// TIA Portal V20 export
// export: Created 2026-10-19T18:01:59.2377084Z, ExportSetting WithDefaults, DisplayName Totally Integrated Automation Portal, DisplayVersion V20 Update 6, DisplayName TIA Portal Openness, DisplayVersion V20 Update 6, DisplayName TIA Portal Version Control Interface, DisplayVersion V20 Update 6, DisplayName SINAMICS Startdrive Advanced, DisplayVersion V20 SP1, DisplayName SINAMICS Startdrive G130, G150, S120, S150, SINAMICS MV, G220, S200, S210, DisplayVersion V20 SP1, DisplayName SINAMICS Startdrive G110M, G120, G120C, G120D, G120P, G115D, DisplayVersion V20 SP1, DisplayName STEP 7 Professional, DisplayVersion V20 Update 6, DisplayName STEP 7 Safety, DisplayVersion V20 Update 2, DisplayName WinCC Basic/Comfort/Advanced, DisplayVersion V20 Update 6, DisplayName WinCC Unified, DisplayVersion V20 Update 6
ORGANIZATION_BLOCK "Main"   // OB1, LAD, ProgramCycle
TITLE = "Main Program Sweep (Cycle)"
{ S7_Optimized_Access := 'TRUE' }
VERSION : 0.1
// stored: AutoNumber true, IsIECCheckEnabled false, SetENOAutomatically false
   VAR_INPUT
      Initial_Call : Bool;   // Initial call of this OB
      Remanence : Bool;   // =True, if remanent data are available
   END_VAR
   VAR_TEMP   // added for the SCL form of the ladder/FBD networks
      _w1 : Bool;
      _w2 : Bool;
      _w3 : Bool;
      _w4 : Bool;
      _w5 : Bool;
   END_VAR
BEGIN

REGION Network 1: Communication
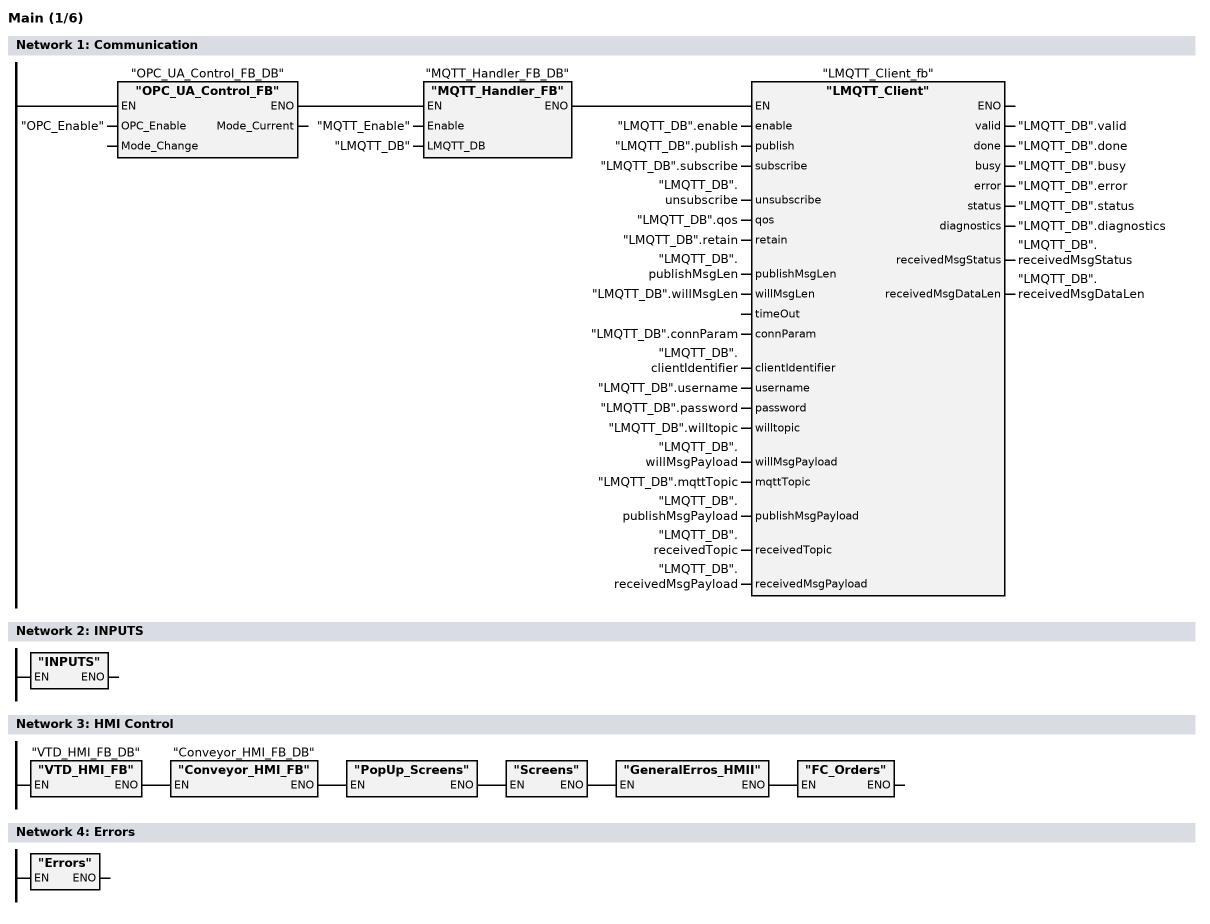
   RUNG wire#powerrail
      "OPC_UA_Control_FB_DB"(OPC_Enable := "OPC_Enable", Mode_Change :=, Mode_Current =>)
      "MQTT_Handler_FB_DB"(Enable := "MQTT_Enable", LMQTT_DB := "LMQTT_DB")
      "LMQTT_Client_fb"(enable := "LMQTT_DB".enable, publish := "LMQTT_DB".publish, subscribe := "LMQTT_DB".subscribe, unsubscribe := "LMQTT_DB".unsubscribe, qos := "LMQTT_DB".qos, retain := "LMQTT_DB".retain, publishMsgLen := "LMQTT_DB".publishMsgLen, willMsgLen := "LMQTT_DB".willMsgLen, timeOut :=, connParam := "LMQTT_DB".connParam, clientIdentifier := "LMQTT_DB".clientIdentifier, username := "LMQTT_DB".username, password := "LMQTT_DB".password, willtopic := "LMQTT_DB".willtopic, willMsgPayload := "LMQTT_DB".willMsgPayload, mqttTopic := "LMQTT_DB".mqttTopic, publishMsgPayload := "LMQTT_DB".publishMsgPayload, receivedTopic := "LMQTT_DB".receivedTopic, receivedMsgPayload := "LMQTT_DB".receivedMsgPayload, valid => "LMQTT_DB".valid, done => "LMQTT_DB".done, busy => "LMQTT_DB".busy, error => "LMQTT_DB".error, status => "LMQTT_DB".status, diagnostics => "LMQTT_DB".diagnostics, receivedMsgStatus => "LMQTT_DB".receivedMsgStatus, receivedMsgDataLen => "LMQTT_DB".receivedMsgDataLen)
   END_RUNG
   // the same network as SCL:
   "OPC_UA_Control_FB_DB"(OPC_Enable := "OPC_Enable", ENO => #_w1);   // "OPC_UA_Control_FB"
   "MQTT_Handler_FB_DB"(EN := #_w1, Enable := "MQTT_Enable", LMQTT_DB := "LMQTT_DB", ENO => #_w2);   // "MQTT_Handler_FB"
   IF #_w2 THEN
       "LMQTT_Client_fb"(enable := "LMQTT_DB".enable,   // "LMQTT_Client"
                         publish := "LMQTT_DB".publish,
                         subscribe := "LMQTT_DB".subscribe,
                         unsubscribe := "LMQTT_DB".unsubscribe,
                         qos := "LMQTT_DB".qos,
                         retain := "LMQTT_DB".retain,
                         publishMsgLen := "LMQTT_DB".publishMsgLen,
                         willMsgLen := "LMQTT_DB".willMsgLen,
                         connParam := "LMQTT_DB".connParam,
                         clientIdentifier := "LMQTT_DB".clientIdentifier,
                         username := "LMQTT_DB".username,
                         password := "LMQTT_DB".password,
                         willtopic := "LMQTT_DB".willtopic,
                         willMsgPayload := "LMQTT_DB".willMsgPayload,
                         mqttTopic := "LMQTT_DB".mqttTopic,
                         publishMsgPayload := "LMQTT_DB".publishMsgPayload,
                         receivedTopic := "LMQTT_DB".receivedTopic,
                         receivedMsgPayload := "LMQTT_DB".receivedMsgPayload,
                         valid => "LMQTT_DB".valid,
                         done => "LMQTT_DB".done,
                         busy => "LMQTT_DB".busy,
                         error => "LMQTT_DB".error,
                         status => "LMQTT_DB".status,
                         diagnostics => "LMQTT_DB".diagnostics,
                         receivedMsgStatus => "LMQTT_DB".receivedMsgStatus,
                         receivedMsgDataLen => "LMQTT_DB".receivedMsgDataLen);
   END_IF;
END_REGION

REGION Network 2: INPUTS
   RUNG wire#powerrail
      "INPUTS"()
   END_RUNG
   // the same network as SCL:
   "INPUTS"();
END_REGION

REGION Network 3: HMI Control
   RUNG wire#powerrail
      "VTD_HMI_FB_DB"()
      "Conveyor_HMI_FB_DB"()
      "PopUp_Screens"()
      "Screens"()
      "GeneralErros_HMII"()
      "FC_Orders"()
   END_RUNG
   // the same network as SCL:
   "VTD_HMI_FB_DB"(ENO => #_w1);   // "VTD_HMI_FB"
   "Conveyor_HMI_FB_DB"(EN := #_w1, ENO => #_w2);   // "Conveyor_HMI_FB"
   "PopUp_Screens"(EN := #_w2, ENO => #_w3);
   "Screens"(EN := #_w3, ENO => #_w4);
   "GeneralErros_HMII"(EN := #_w4, ENO => #_w5);
   IF #_w5 THEN "FC_Orders"(); END_IF;
END_REGION

REGION Network 4: Errors
   RUNG wire#powerrail
      "Errors"()
   END_RUNG
   // the same network as SCL:
   "Errors"();
END_REGION

REGION Network 5: Carousel Conveyors
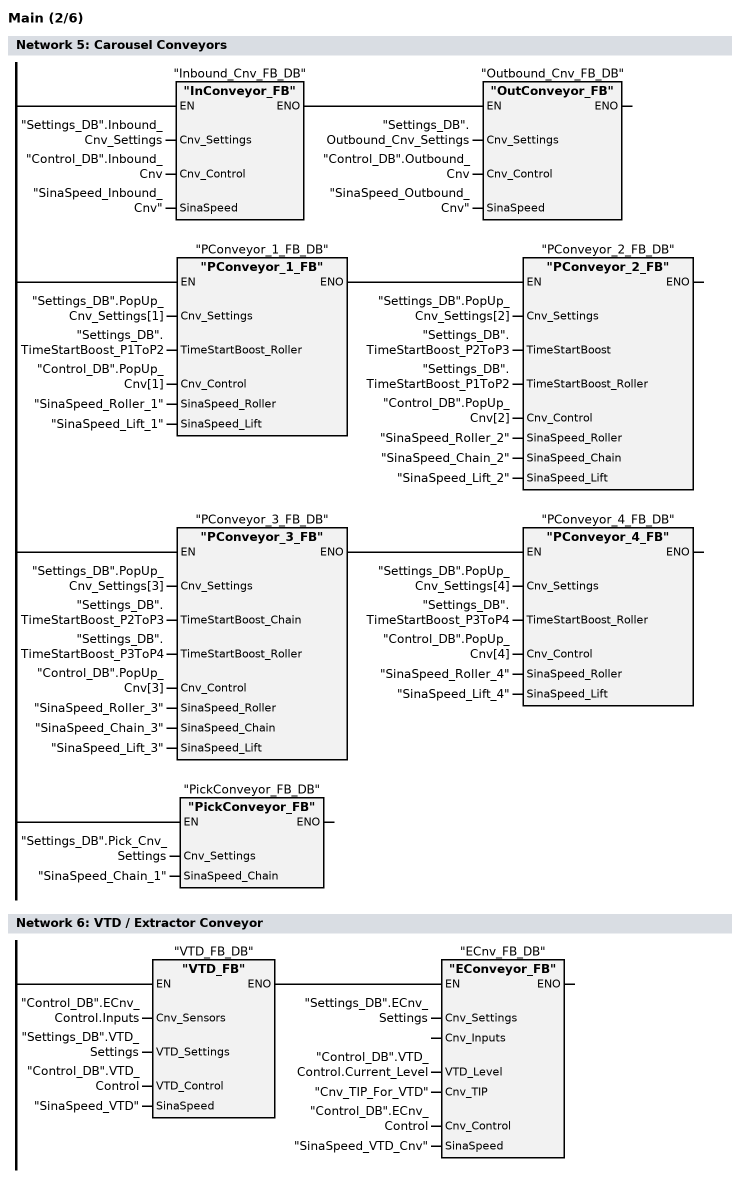
   RUNG wire#powerrail
      "Inbound_Cnv_FB_DB"(Cnv_Settings := "Settings_DB".Inbound_Cnv_Settings, Cnv_Control := "Control_DB".Inbound_Cnv, SinaSpeed := "SinaSpeed_Inbound_Cnv")
      "Outbound_Cnv_FB_DB"(Cnv_Settings := "Settings_DB".Outbound_Cnv_Settings, Cnv_Control := "Control_DB".Outbound_Cnv, SinaSpeed := "SinaSpeed_Outbound_Cnv")
   END_RUNG
   RUNG wire#powerrail
      "PConveyor_1_FB_DB"(Cnv_Settings := "Settings_DB".PopUp_Cnv_Settings[1], TimeStartBoost_Roller := "Settings_DB".TimeStartBoost_P1ToP2, Cnv_Control := "Control_DB".PopUp_Cnv[1], SinaSpeed_Roller := "SinaSpeed_Roller_1", SinaSpeed_Lift := "SinaSpeed_Lift_1")
      "PConveyor_2_FB_DB"(Cnv_Settings := "Settings_DB".PopUp_Cnv_Settings[2], TimeStartBoost := "Settings_DB".TimeStartBoost_P2ToP3, TimeStartBoost_Roller := "Settings_DB".TimeStartBoost_P1ToP2, Cnv_Control := "Control_DB".PopUp_Cnv[2], SinaSpeed_Roller := "SinaSpeed_Roller_2", SinaSpeed_Chain := "SinaSpeed_Chain_2", SinaSpeed_Lift := "SinaSpeed_Lift_2")
   END_RUNG
   RUNG wire#powerrail
      "PConveyor_3_FB_DB"(Cnv_Settings := "Settings_DB".PopUp_Cnv_Settings[3], TimeStartBoost_Chain := "Settings_DB".TimeStartBoost_P2ToP3, TimeStartBoost_Roller := "Settings_DB".TimeStartBoost_P3ToP4, Cnv_Control := "Control_DB".PopUp_Cnv[3], SinaSpeed_Roller := "SinaSpeed_Roller_3", SinaSpeed_Chain := "SinaSpeed_Chain_3", SinaSpeed_Lift := "SinaSpeed_Lift_3")
      "PConveyor_4_FB_DB"(Cnv_Settings := "Settings_DB".PopUp_Cnv_Settings[4], TimeStartBoost_Roller := "Settings_DB".TimeStartBoost_P3ToP4, Cnv_Control := "Control_DB".PopUp_Cnv[4], SinaSpeed_Roller := "SinaSpeed_Roller_4", SinaSpeed_Lift := "SinaSpeed_Lift_4")
   END_RUNG
   RUNG wire#powerrail
      "PickConveyor_FB_DB"(Cnv_Settings := "Settings_DB".Pick_Cnv_Settings, SinaSpeed_Chain := "SinaSpeed_Chain_1")
   END_RUNG
   // the same network as SCL:
   "Inbound_Cnv_FB_DB"(Cnv_Settings := "Settings_DB".Inbound_Cnv_Settings,   // "InConveyor_FB"
                       Cnv_Control := "Control_DB".Inbound_Cnv,
                       SinaSpeed := "SinaSpeed_Inbound_Cnv",
                       ENO => #_w1);
   IF #_w1 THEN
       "Outbound_Cnv_FB_DB"(Cnv_Settings := "Settings_DB".Outbound_Cnv_Settings,   // "OutConveyor_FB"
                            Cnv_Control := "Control_DB".Outbound_Cnv,
                            SinaSpeed := "SinaSpeed_Outbound_Cnv");
   END_IF;
   "PConveyor_1_FB_DB"(Cnv_Settings := "Settings_DB".PopUp_Cnv_Settings[1],   // "PConveyor_1_FB"
                       TimeStartBoost_Roller := "Settings_DB".TimeStartBoost_P1ToP2,
                       Cnv_Control := "Control_DB".PopUp_Cnv[1],
                       SinaSpeed_Roller := "SinaSpeed_Roller_1",
                       SinaSpeed_Lift := "SinaSpeed_Lift_1",
                       ENO => #_w2);
   IF #_w2 THEN
       "PConveyor_2_FB_DB"(Cnv_Settings := "Settings_DB".PopUp_Cnv_Settings[2],   // "PConveyor_2_FB"
                           TimeStartBoost := "Settings_DB".TimeStartBoost_P2ToP3,
                           TimeStartBoost_Roller := "Settings_DB".TimeStartBoost_P1ToP2,
                           Cnv_Control := "Control_DB".PopUp_Cnv[2],
                           SinaSpeed_Roller := "SinaSpeed_Roller_2",
                           SinaSpeed_Chain := "SinaSpeed_Chain_2",
                           SinaSpeed_Lift := "SinaSpeed_Lift_2");
   END_IF;
   "PConveyor_3_FB_DB"(Cnv_Settings := "Settings_DB".PopUp_Cnv_Settings[3],   // "PConveyor_3_FB"
                       TimeStartBoost_Chain := "Settings_DB".TimeStartBoost_P2ToP3,
                       TimeStartBoost_Roller := "Settings_DB".TimeStartBoost_P3ToP4,
                       Cnv_Control := "Control_DB".PopUp_Cnv[3],
                       SinaSpeed_Roller := "SinaSpeed_Roller_3",
                       SinaSpeed_Chain := "SinaSpeed_Chain_3",
                       SinaSpeed_Lift := "SinaSpeed_Lift_3",
                       ENO => #_w3);
   IF #_w3 THEN
       "PConveyor_4_FB_DB"(Cnv_Settings := "Settings_DB".PopUp_Cnv_Settings[4],   // "PConveyor_4_FB"
                           TimeStartBoost_Roller := "Settings_DB".TimeStartBoost_P3ToP4,
                           Cnv_Control := "Control_DB".PopUp_Cnv[4],
                           SinaSpeed_Roller := "SinaSpeed_Roller_4",
                           SinaSpeed_Lift := "SinaSpeed_Lift_4");
   END_IF;
   "PickConveyor_FB_DB"(Cnv_Settings := "Settings_DB".Pick_Cnv_Settings, SinaSpeed_Chain := "SinaSpeed_Chain_1");   // "PickConveyor_FB"
END_REGION

REGION Network 6: VTD / Extractor Conveyor
   RUNG wire#powerrail
      "VTD_FB_DB"(Cnv_Sensors := "Control_DB".ECnv_Control.Inputs, VTD_Settings := "Settings_DB".VTD_Settings, VTD_Control := "Control_DB".VTD_Control, SinaSpeed := "SinaSpeed_VTD")
      "ECnv_FB_DB"(Cnv_Settings := "Settings_DB".ECnv_Settings, Cnv_Inputs :=, VTD_Level := "Control_DB".VTD_Control.Current_Level, Cnv_TIP := "Cnv_TIP_For_VTD", Cnv_Control := "Control_DB".ECnv_Control, SinaSpeed := "SinaSpeed_VTD_Cnv")
   END_RUNG
   // the same network as SCL:
   "VTD_FB_DB"(Cnv_Sensors := "Control_DB".ECnv_Control.Inputs,   // "VTD_FB"
               VTD_Settings := "Settings_DB".VTD_Settings,
               VTD_Control := "Control_DB".VTD_Control,
               SinaSpeed := "SinaSpeed_VTD",
               ENO => #_w1);
   IF #_w1 THEN
       "ECnv_FB_DB"(Cnv_Settings := "Settings_DB".ECnv_Settings,   // "EConveyor_FB"
                    VTD_Level := "Control_DB".VTD_Control.Current_Level,
                    Cnv_TIP := "Cnv_TIP_For_VTD",
                    Cnv_Control := "Control_DB".ECnv_Control,
                    SinaSpeed := "SinaSpeed_VTD_Cnv");
   END_IF;
END_REGION

REGION Network 7: Level Conveyors
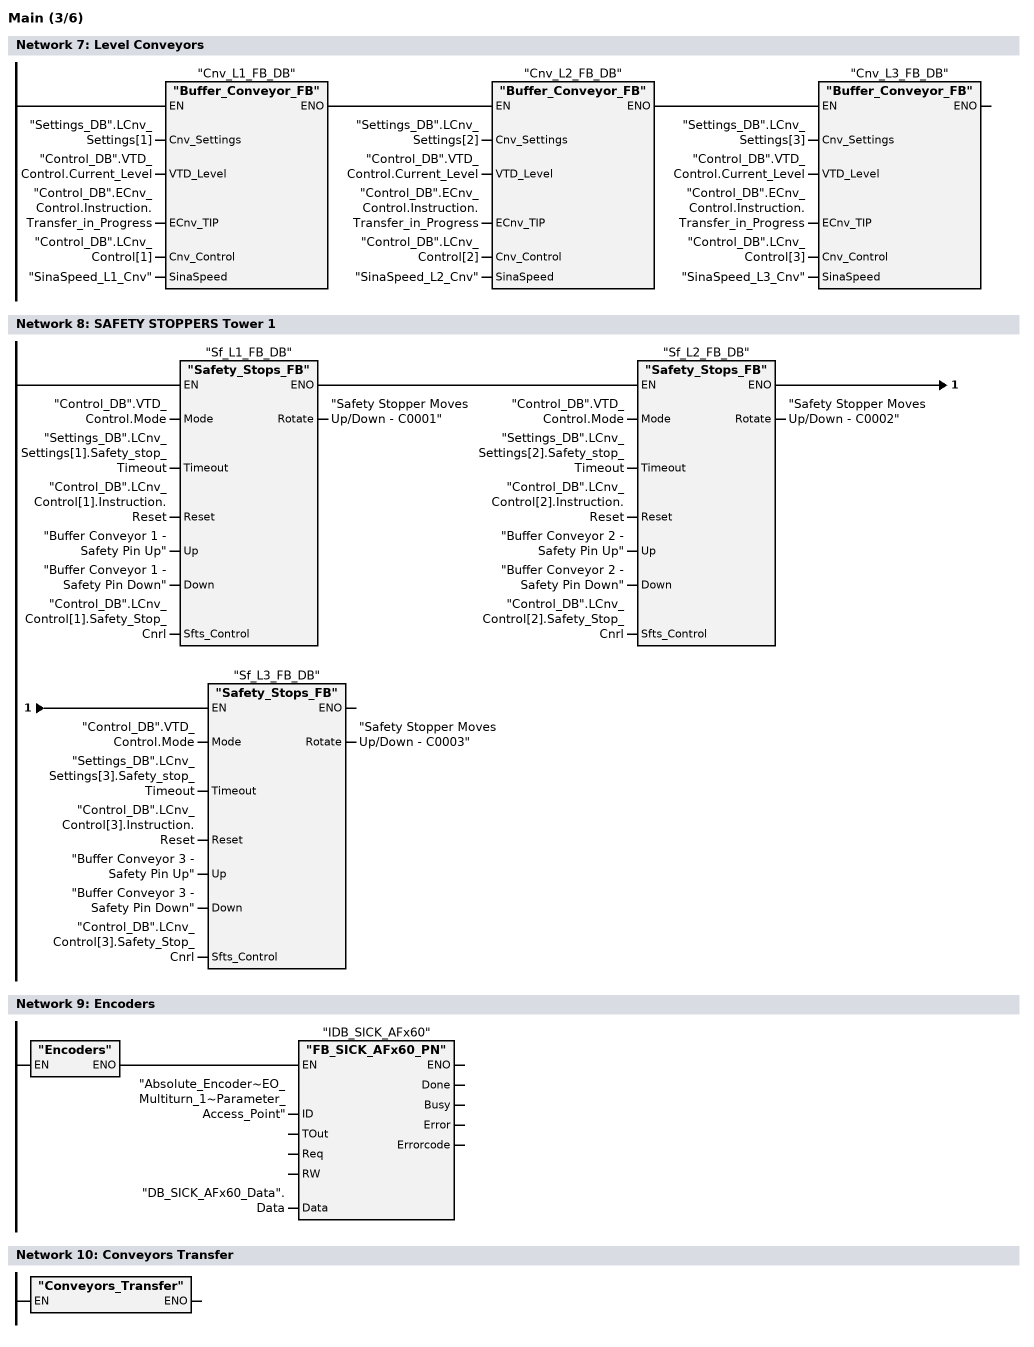
   RUNG wire#powerrail
      "Cnv_L1_FB_DB"(Cnv_Settings := "Settings_DB".LCnv_Settings[1], VTD_Level := "Control_DB".VTD_Control.Current_Level, ECnv_TIP := "Control_DB".ECnv_Control.Instruction.Transfer_in_Progress, Cnv_Control := "Control_DB".LCnv_Control[1], SinaSpeed := "SinaSpeed_L1_Cnv")
      "Cnv_L2_FB_DB"(Cnv_Settings := "Settings_DB".LCnv_Settings[2], VTD_Level := "Control_DB".VTD_Control.Current_Level, ECnv_TIP := "Control_DB".ECnv_Control.Instruction.Transfer_in_Progress, Cnv_Control := "Control_DB".LCnv_Control[2], SinaSpeed := "SinaSpeed_L2_Cnv")
      "Cnv_L3_FB_DB"(Cnv_Settings := "Settings_DB".LCnv_Settings[3], VTD_Level := "Control_DB".VTD_Control.Current_Level, ECnv_TIP := "Control_DB".ECnv_Control.Instruction.Transfer_in_Progress, Cnv_Control := "Control_DB".LCnv_Control[3], SinaSpeed := "SinaSpeed_L3_Cnv")
   END_RUNG
   // the same network as SCL:
   "Cnv_L1_FB_DB"(Cnv_Settings := "Settings_DB".LCnv_Settings[1],   // "Buffer_Conveyor_FB"
                  VTD_Level := "Control_DB".VTD_Control.Current_Level,
                  ECnv_TIP := "Control_DB".ECnv_Control.Instruction.Transfer_in_Progress,
                  Cnv_Control := "Control_DB".LCnv_Control[1],
                  SinaSpeed := "SinaSpeed_L1_Cnv",
                  ENO => #_w1);
   "Cnv_L2_FB_DB"(EN := #_w1,   // "Buffer_Conveyor_FB"
                  Cnv_Settings := "Settings_DB".LCnv_Settings[2],
                  VTD_Level := "Control_DB".VTD_Control.Current_Level,
                  ECnv_TIP := "Control_DB".ECnv_Control.Instruction.Transfer_in_Progress,
                  Cnv_Control := "Control_DB".LCnv_Control[2],
                  SinaSpeed := "SinaSpeed_L2_Cnv",
                  ENO => #_w2);
   IF #_w2 THEN
       "Cnv_L3_FB_DB"(Cnv_Settings := "Settings_DB".LCnv_Settings[3],   // "Buffer_Conveyor_FB"
                      VTD_Level := "Control_DB".VTD_Control.Current_Level,
                      ECnv_TIP := "Control_DB".ECnv_Control.Instruction.Transfer_in_Progress,
                      Cnv_Control := "Control_DB".LCnv_Control[3],
                      SinaSpeed := "SinaSpeed_L3_Cnv");
   END_IF;
END_REGION

REGION Network 8: SAFETY STOPPERS Tower 1
   RUNG wire#powerrail
      "Sf_L1_FB_DB"(Mode := "Control_DB".VTD_Control.Mode, Timeout := "Settings_DB".LCnv_Settings[1].Safety_stop_Timeout, Reset := "Control_DB".LCnv_Control[1].Instruction.Reset, Up := "Buffer Conveyor 1 - Safety Pin Up", Down := "Buffer Conveyor 1 - Safety Pin Down", Sfts_Control := "Control_DB".LCnv_Control[1].Safety_Stop_Cnrl, Rotate => "Safety Stopper Moves Up/Down - C0001")
      "Sf_L2_FB_DB"(Mode := "Control_DB".VTD_Control.Mode, Timeout := "Settings_DB".LCnv_Settings[2].Safety_stop_Timeout, Reset := "Control_DB".LCnv_Control[2].Instruction.Reset, Up := "Buffer Conveyor 2 - Safety Pin Up", Down := "Buffer Conveyor 2 - Safety Pin Down", Sfts_Control := "Control_DB".LCnv_Control[2].Safety_Stop_Cnrl, Rotate => "Safety Stopper Moves Up/Down - C0002")
      "Sf_L3_FB_DB"(Mode := "Control_DB".VTD_Control.Mode, Timeout := "Settings_DB".LCnv_Settings[3].Safety_stop_Timeout, Reset := "Control_DB".LCnv_Control[3].Instruction.Reset, Up := "Buffer Conveyor 3 - Safety Pin Up", Down := "Buffer Conveyor 3 - Safety Pin Down", Sfts_Control := "Control_DB".LCnv_Control[3].Safety_Stop_Cnrl, Rotate => "Safety Stopper Moves Up/Down - C0003")
   END_RUNG
   // the same network as SCL:
   "Sf_L1_FB_DB"(Mode := "Control_DB".VTD_Control.Mode,   // "Safety_Stops_FB"
                 Timeout := "Settings_DB".LCnv_Settings[1].Safety_stop_Timeout,
                 Reset := "Control_DB".LCnv_Control[1].Instruction.Reset,
                 Up := "Buffer Conveyor 1 - Safety Pin Up",
                 Down := "Buffer Conveyor 1 - Safety Pin Down",
                 Sfts_Control := "Control_DB".LCnv_Control[1].Safety_Stop_Cnrl,
                 Rotate => "Safety Stopper Moves Up/Down - C0001",
                 ENO => #_w1);
   "Sf_L2_FB_DB"(EN := #_w1,   // "Safety_Stops_FB"
                 Mode := "Control_DB".VTD_Control.Mode,
                 Timeout := "Settings_DB".LCnv_Settings[2].Safety_stop_Timeout,
                 Reset := "Control_DB".LCnv_Control[2].Instruction.Reset,
                 Up := "Buffer Conveyor 2 - Safety Pin Up",
                 Down := "Buffer Conveyor 2 - Safety Pin Down",
                 Sfts_Control := "Control_DB".LCnv_Control[2].Safety_Stop_Cnrl,
                 Rotate => "Safety Stopper Moves Up/Down - C0002",
                 ENO => #_w2);
   IF #_w2 THEN
       "Sf_L3_FB_DB"(Mode := "Control_DB".VTD_Control.Mode,   // "Safety_Stops_FB"
                     Timeout := "Settings_DB".LCnv_Settings[3].Safety_stop_Timeout,
                     Reset := "Control_DB".LCnv_Control[3].Instruction.Reset,
                     Up := "Buffer Conveyor 3 - Safety Pin Up",
                     Down := "Buffer Conveyor 3 - Safety Pin Down",
                     Sfts_Control := "Control_DB".LCnv_Control[3].Safety_Stop_Cnrl,
                     Rotate => "Safety Stopper Moves Up/Down - C0003");
   END_IF;
END_REGION

REGION Network 9: Encoders
   RUNG wire#powerrail
      "Encoders"()
      "IDB_SICK_AFx60"(ID := "Absolute_Encoder~EO_Multiturn_1~Parameter_Access_Point", TOut :=, Req :=, RW :=, Data := "DB_SICK_AFx60_Data".Data, Done =>, Busy =>, Error =>, Errorcode =>)
   END_RUNG
   // the same network as SCL:
   "Encoders"(ENO => #_w1);
   IF #_w1 THEN
       "IDB_SICK_AFx60"(ID := "Absolute_Encoder~EO_Multiturn_1~Parameter_Access_Point",   // "FB_SICK_AFx60_PN"
                        Data := "DB_SICK_AFx60_Data".Data);
   END_IF;
END_REGION

REGION Network 10: Conveyors Transfer
   RUNG wire#powerrail
      "Conveyors_Transfer"()
   END_RUNG
   // the same network as SCL:
   "Conveyors_Transfer"();
END_REGION

REGION Network 11: Lightbar
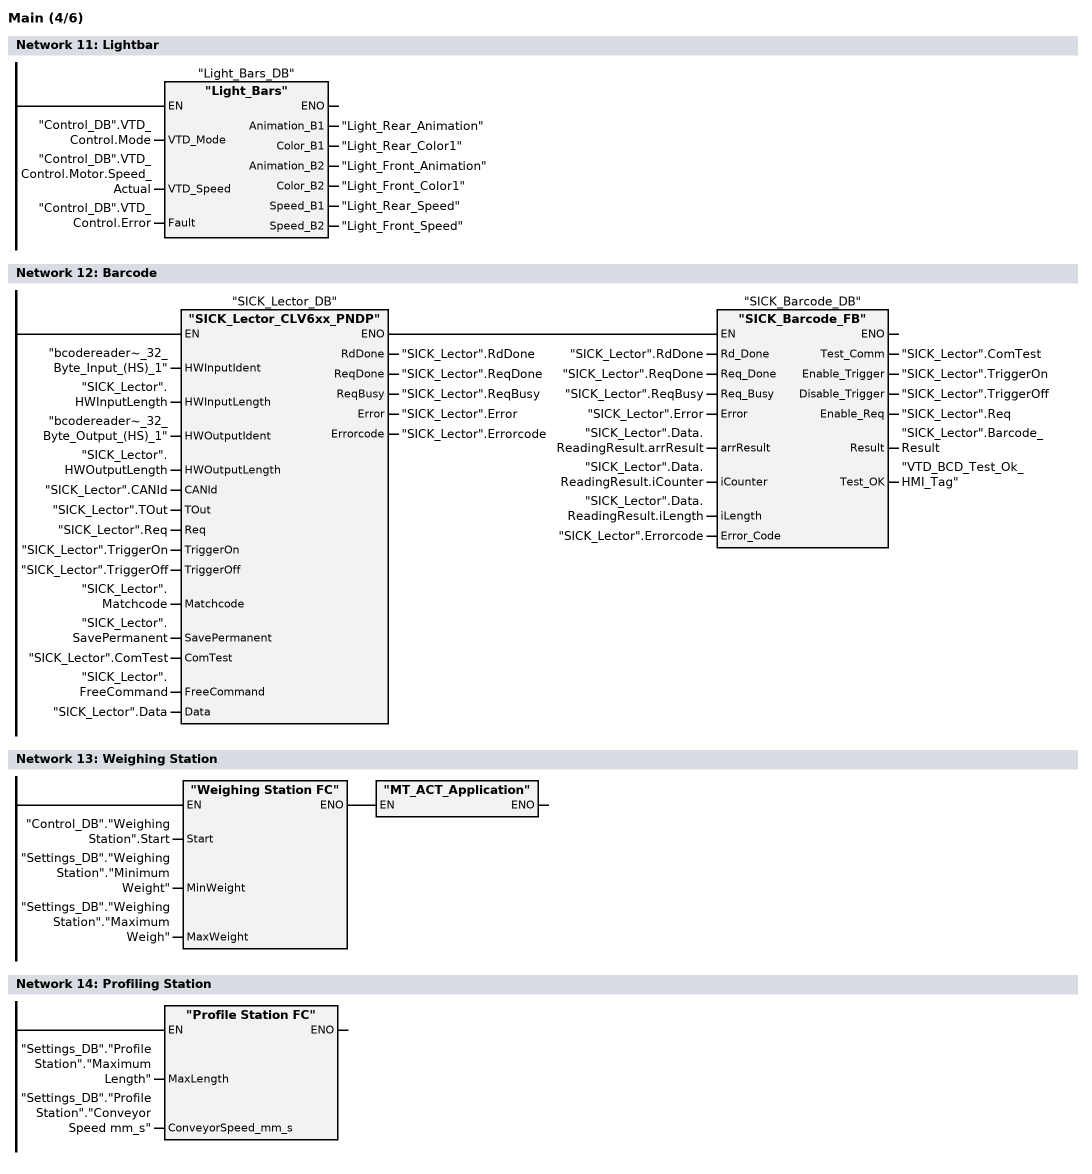
   RUNG wire#powerrail
      "Light_Bars_DB"(VTD_Mode := "Control_DB".VTD_Control.Mode, VTD_Speed := "Control_DB".VTD_Control.Motor.Speed_Actual, Fault := "Control_DB".VTD_Control.Error, Animation_B1 => "Light_Rear_Animation", Color_B1 => "Light_Rear_Color1", Animation_B2 => "Light_Front_Animation", Color_B2 => "Light_Front_Color1", Speed_B1 => "Light_Rear_Speed", Speed_B2 => "Light_Front_Speed")
   END_RUNG
   // the same network as SCL:
   "Light_Bars_DB"(VTD_Mode := "Control_DB".VTD_Control.Mode,   // "Light_Bars"
                   VTD_Speed := "Control_DB".VTD_Control.Motor.Speed_Actual,
                   Fault := "Control_DB".VTD_Control.Error,
                   Animation_B1 => "Light_Rear_Animation",
                   Color_B1 => "Light_Rear_Color1",
                   Animation_B2 => "Light_Front_Animation",
                   Color_B2 => "Light_Front_Color1",
                   Speed_B1 => "Light_Rear_Speed",
                   Speed_B2 => "Light_Front_Speed");
END_REGION

REGION Network 12: Barcode
   RUNG wire#powerrail
      "SICK_Lector_DB"(HWInputIdent := "bcodereader~_32_Byte_Input_(HS)_1", HWInputLength := "SICK_Lector".HWInputLength, HWOutputIdent := "bcodereader~_32_Byte_Output_(HS)_1", HWOutputLength := "SICK_Lector".HWOutputLength, CANId := "SICK_Lector".CANId, TOut := "SICK_Lector".TOut, Req := "SICK_Lector".Req, TriggerOn := "SICK_Lector".TriggerOn, TriggerOff := "SICK_Lector".TriggerOff, Matchcode := "SICK_Lector".Matchcode, SavePermanent := "SICK_Lector".SavePermanent, ComTest := "SICK_Lector".ComTest, FreeCommand := "SICK_Lector".FreeCommand, Data := "SICK_Lector".Data, RdDone => "SICK_Lector".RdDone, ReqDone => "SICK_Lector".ReqDone, ReqBusy => "SICK_Lector".ReqBusy, Error => "SICK_Lector".Error, Errorcode => "SICK_Lector".Errorcode)
      "SICK_Barcode_DB"(Rd_Done := "SICK_Lector".RdDone, Req_Done := "SICK_Lector".ReqDone, Req_Busy := "SICK_Lector".ReqBusy, Error := "SICK_Lector".Error, arrResult := "SICK_Lector".Data.ReadingResult.arrResult, iCounter := "SICK_Lector".Data.ReadingResult.iCounter, iLength := "SICK_Lector".Data.ReadingResult.iLength, Error_Code := "SICK_Lector".Errorcode, Test_Comm => "SICK_Lector".ComTest, Enable_Trigger => "SICK_Lector".TriggerOn, Disable_Trigger => "SICK_Lector".TriggerOff, Enable_Req => "SICK_Lector".Req, Result => "SICK_Lector".Barcode_Result, Test_OK => "VTD_BCD_Test_Ok_HMI_Tag")
   END_RUNG
   // the same network as SCL:
   "SICK_Lector_DB"(HWInputIdent := "bcodereader~_32_Byte_Input_(HS)_1",   // "SICK_Lector_CLV6xx_PNDP"
                    HWInputLength := "SICK_Lector".HWInputLength,
                    HWOutputIdent := "bcodereader~_32_Byte_Output_(HS)_1",
                    HWOutputLength := "SICK_Lector".HWOutputLength,
                    CANId := "SICK_Lector".CANId,
                    TOut := "SICK_Lector".TOut,
                    Req := "SICK_Lector".Req,
                    TriggerOn := "SICK_Lector".TriggerOn,
                    TriggerOff := "SICK_Lector".TriggerOff,
                    Matchcode := "SICK_Lector".Matchcode,
                    SavePermanent := "SICK_Lector".SavePermanent,
                    ComTest := "SICK_Lector".ComTest,
                    FreeCommand := "SICK_Lector".FreeCommand,
                    Data := "SICK_Lector".Data,
                    RdDone => "SICK_Lector".RdDone,
                    ReqDone => "SICK_Lector".ReqDone,
                    ReqBusy => "SICK_Lector".ReqBusy,
                    Error => "SICK_Lector".Error,
                    Errorcode => "SICK_Lector".Errorcode,
                    ENO => #_w1);
   IF #_w1 THEN
       "SICK_Barcode_DB"(Rd_Done := "SICK_Lector".RdDone,   // "SICK_Barcode_FB"
                         Req_Done := "SICK_Lector".ReqDone,
                         Req_Busy := "SICK_Lector".ReqBusy,
                         Error := "SICK_Lector".Error,
                         arrResult := "SICK_Lector".Data.ReadingResult.arrResult,
                         iCounter := "SICK_Lector".Data.ReadingResult.iCounter,
                         iLength := "SICK_Lector".Data.ReadingResult.iLength,
                         Error_Code := "SICK_Lector".Errorcode,
                         Test_Comm => "SICK_Lector".ComTest,
                         Enable_Trigger => "SICK_Lector".TriggerOn,
                         Disable_Trigger => "SICK_Lector".TriggerOff,
                         Enable_Req => "SICK_Lector".Req,
                         Result => "SICK_Lector".Barcode_Result,
                         Test_OK => "VTD_BCD_Test_Ok_HMI_Tag");
   END_IF;
END_REGION

REGION Network 13: Weighing Station
   RUNG wire#powerrail
      "Weighing Station FC"(Start := "Control_DB"."Weighing Station".Start, MinWeight := "Settings_DB"."Weighing Station"."Minimum Weight", MaxWeight := "Settings_DB"."Weighing Station"."Maximum Weigh")
      "MT_ACT_Application"()
   END_RUNG
   // the same network as SCL:
   "Weighing Station FC"(Start := "Control_DB"."Weighing Station".Start,
                         MinWeight := "Settings_DB"."Weighing Station"."Minimum Weight",
                         MaxWeight := "Settings_DB"."Weighing Station"."Maximum Weigh",
                         ENO => #_w1);
   IF #_w1 THEN "MT_ACT_Application"(); END_IF;
END_REGION

REGION Network 14: Profiling Station
   RUNG wire#powerrail
      "Profile Station FC"(MaxLength := "Settings_DB"."Profile Station"."Maximum Length", ConveyorSpeed_mm_s := "Settings_DB"."Profile Station"."Conveyor Speed mm_s")
   END_RUNG
   // the same network as SCL:
   "Profile Station FC"(MaxLength := "Settings_DB"."Profile Station"."Maximum Length",
                        ConveyorSpeed_mm_s := "Settings_DB"."Profile Station"."Conveyor Speed mm_s");
END_REGION

REGION Network 15: Barcode Stations
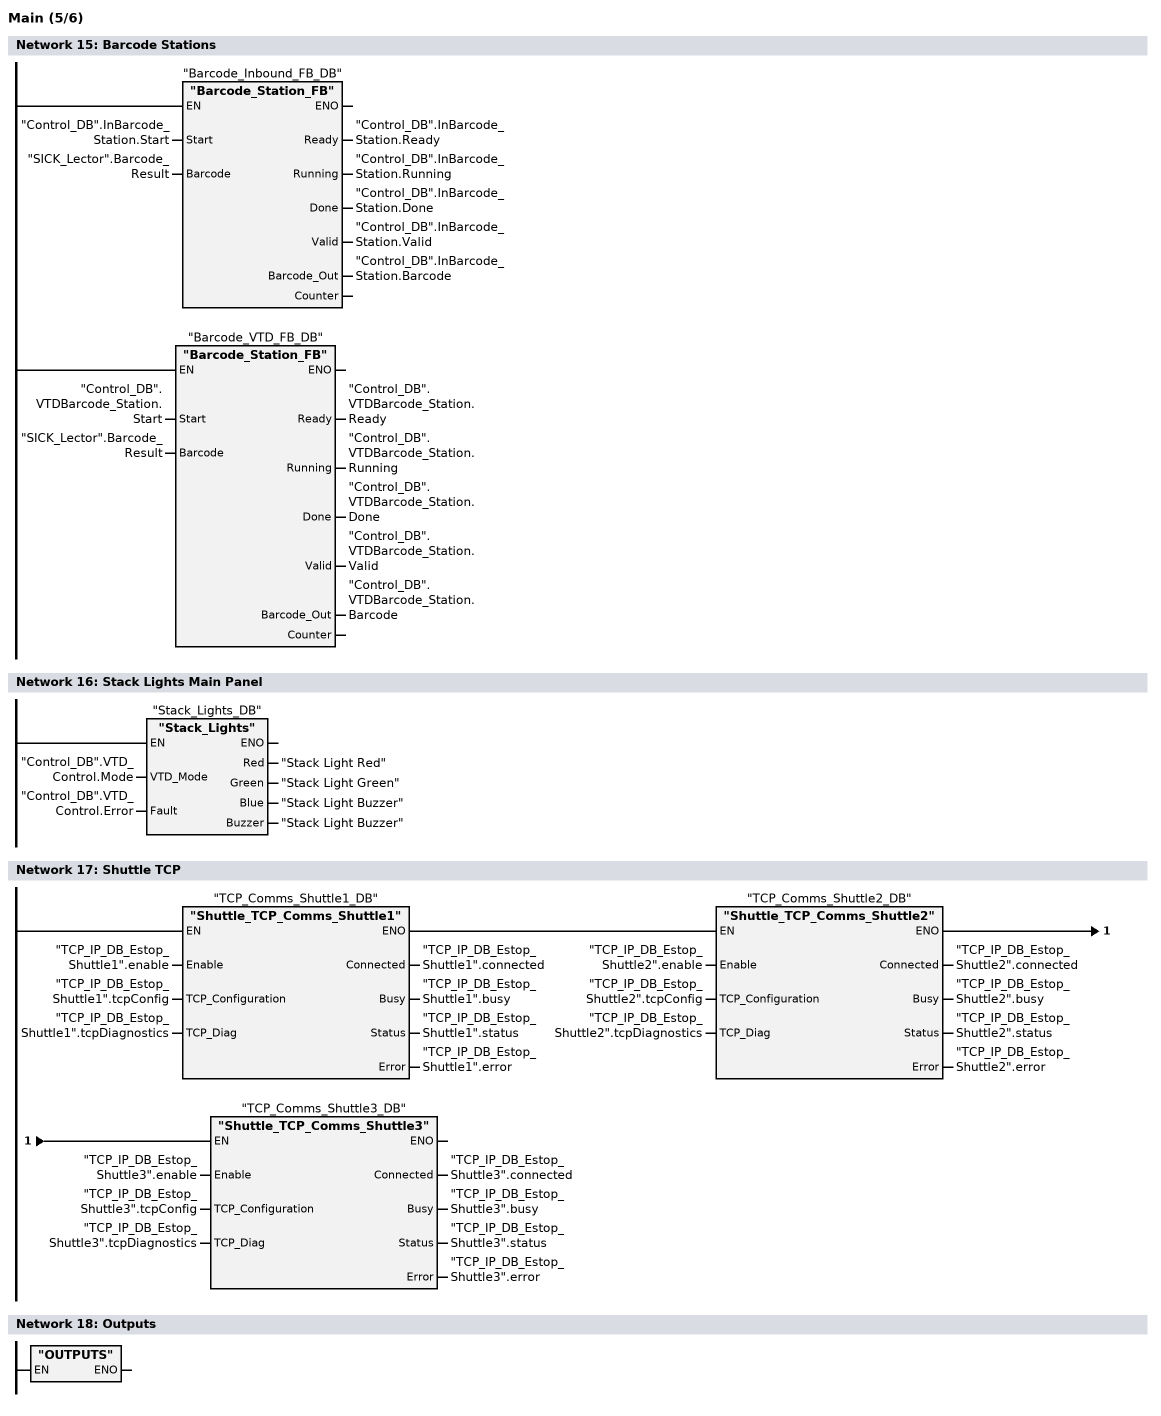
   RUNG wire#powerrail
      "Barcode_Inbound_FB_DB"(Start := "Control_DB".InBarcode_Station.Start, Barcode := "SICK_Lector".Barcode_Result, Ready => "Control_DB".InBarcode_Station.Ready, Running => "Control_DB".InBarcode_Station.Running, Done => "Control_DB".InBarcode_Station.Done, Valid => "Control_DB".InBarcode_Station.Valid, Barcode_Out => "Control_DB".InBarcode_Station.Barcode, "Counter" =>)
   END_RUNG
   RUNG wire#powerrail
      "Barcode_VTD_FB_DB"(Start := "Control_DB".VTDBarcode_Station.Start, Barcode := "SICK_Lector".Barcode_Result, Ready => "Control_DB".VTDBarcode_Station.Ready, Running => "Control_DB".VTDBarcode_Station.Running, Done => "Control_DB".VTDBarcode_Station.Done, Valid => "Control_DB".VTDBarcode_Station.Valid, Barcode_Out => "Control_DB".VTDBarcode_Station.Barcode, "Counter" =>)
   END_RUNG
   // the same network as SCL:
   "Barcode_Inbound_FB_DB"(Start := "Control_DB".InBarcode_Station.Start,   // "Barcode_Station_FB"
                           Barcode := "SICK_Lector".Barcode_Result,
                           Ready => "Control_DB".InBarcode_Station.Ready,
                           Running => "Control_DB".InBarcode_Station.Running,
                           Done => "Control_DB".InBarcode_Station.Done,
                           Valid => "Control_DB".InBarcode_Station.Valid,
                           Barcode_Out => "Control_DB".InBarcode_Station.Barcode);
   "Barcode_VTD_FB_DB"(Start := "Control_DB".VTDBarcode_Station.Start,   // "Barcode_Station_FB"
                       Barcode := "SICK_Lector".Barcode_Result,
                       Ready => "Control_DB".VTDBarcode_Station.Ready,
                       Running => "Control_DB".VTDBarcode_Station.Running,
                       Done => "Control_DB".VTDBarcode_Station.Done,
                       Valid => "Control_DB".VTDBarcode_Station.Valid,
                       Barcode_Out => "Control_DB".VTDBarcode_Station.Barcode);
END_REGION

REGION Network 16: Stack Lights Main Panel
   RUNG wire#powerrail
      "Stack_Lights_DB"(VTD_Mode := "Control_DB".VTD_Control.Mode, Fault := "Control_DB".VTD_Control.Error, Red => "Stack Light Red", Green => "Stack Light Green", Blue => "Stack Light Buzzer", Buzzer => "Stack Light Buzzer")
   END_RUNG
   // the same network as SCL:
   "Stack_Lights_DB"(VTD_Mode := "Control_DB".VTD_Control.Mode,   // "Stack_Lights"
                     Fault := "Control_DB".VTD_Control.Error,
                     Red => "Stack Light Red",
                     Green => "Stack Light Green",
                     Blue => "Stack Light Buzzer",
                     Buzzer => "Stack Light Buzzer");
END_REGION

REGION Network 17: Shuttle TCP
   RUNG wire#powerrail
      "TCP_Comms_Shuttle1_DB"(Enable := "TCP_IP_DB_Estop_Shuttle1".enable, TCP_Configuration := "TCP_IP_DB_Estop_Shuttle1".tcpConfig, TCP_Diag := "TCP_IP_DB_Estop_Shuttle1".tcpDiagnostics, Connected => "TCP_IP_DB_Estop_Shuttle1".connected, Busy => "TCP_IP_DB_Estop_Shuttle1".busy, Status => "TCP_IP_DB_Estop_Shuttle1".status, Error => "TCP_IP_DB_Estop_Shuttle1".error)
      "TCP_Comms_Shuttle2_DB"(Enable := "TCP_IP_DB_Estop_Shuttle2".enable, TCP_Configuration := "TCP_IP_DB_Estop_Shuttle2".tcpConfig, TCP_Diag := "TCP_IP_DB_Estop_Shuttle2".tcpDiagnostics, Connected => "TCP_IP_DB_Estop_Shuttle2".connected, Busy => "TCP_IP_DB_Estop_Shuttle2".busy, Status => "TCP_IP_DB_Estop_Shuttle2".status, Error => "TCP_IP_DB_Estop_Shuttle2".error)
      "TCP_Comms_Shuttle3_DB"(Enable := "TCP_IP_DB_Estop_Shuttle3".enable, TCP_Configuration := "TCP_IP_DB_Estop_Shuttle3".tcpConfig, TCP_Diag := "TCP_IP_DB_Estop_Shuttle3".tcpDiagnostics, Connected => "TCP_IP_DB_Estop_Shuttle3".connected, Busy => "TCP_IP_DB_Estop_Shuttle3".busy, Status => "TCP_IP_DB_Estop_Shuttle3".status, Error => "TCP_IP_DB_Estop_Shuttle3".error)
   END_RUNG
   // the same network as SCL:
   "TCP_Comms_Shuttle1_DB"(Enable := "TCP_IP_DB_Estop_Shuttle1".enable,   // "Shuttle_TCP_Comms_Shuttle1"
                           TCP_Configuration := "TCP_IP_DB_Estop_Shuttle1".tcpConfig,
                           TCP_Diag := "TCP_IP_DB_Estop_Shuttle1".tcpDiagnostics,
                           Connected => "TCP_IP_DB_Estop_Shuttle1".connected,
                           Busy => "TCP_IP_DB_Estop_Shuttle1".busy,
                           Status => "TCP_IP_DB_Estop_Shuttle1".status,
                           Error => "TCP_IP_DB_Estop_Shuttle1".error,
                           ENO => #_w1);
   "TCP_Comms_Shuttle2_DB"(EN := #_w1,   // "Shuttle_TCP_Comms_Shuttle2"
                           Enable := "TCP_IP_DB_Estop_Shuttle2".enable,
                           TCP_Configuration := "TCP_IP_DB_Estop_Shuttle2".tcpConfig,
                           TCP_Diag := "TCP_IP_DB_Estop_Shuttle2".tcpDiagnostics,
                           Connected => "TCP_IP_DB_Estop_Shuttle2".connected,
                           Busy => "TCP_IP_DB_Estop_Shuttle2".busy,
                           Status => "TCP_IP_DB_Estop_Shuttle2".status,
                           Error => "TCP_IP_DB_Estop_Shuttle2".error,
                           ENO => #_w2);
   IF #_w2 THEN
       "TCP_Comms_Shuttle3_DB"(Enable := "TCP_IP_DB_Estop_Shuttle3".enable,   // "Shuttle_TCP_Comms_Shuttle3"
                               TCP_Configuration := "TCP_IP_DB_Estop_Shuttle3".tcpConfig,
                               TCP_Diag := "TCP_IP_DB_Estop_Shuttle3".tcpDiagnostics,
                               Connected => "TCP_IP_DB_Estop_Shuttle3".connected,
                               Busy => "TCP_IP_DB_Estop_Shuttle3".busy,
                               Status => "TCP_IP_DB_Estop_Shuttle3".status,
                               Error => "TCP_IP_DB_Estop_Shuttle3".error);
   END_IF;
END_REGION

REGION Network 18: Outputs
   RUNG wire#powerrail
      "OUTPUTS"()
   END_RUNG
   // the same network as SCL:
   "OUTPUTS"();
END_REGION

REGION Network 19: System Order Table - Carousel
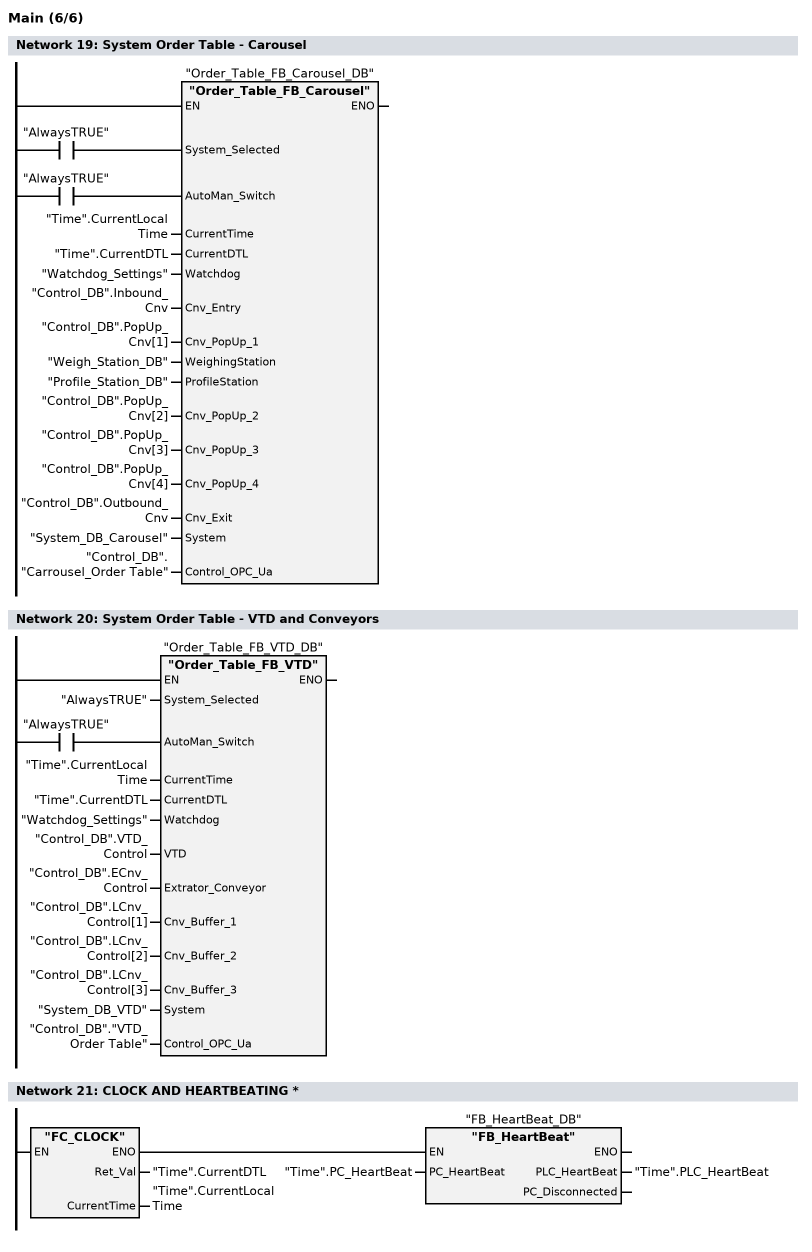
   RUNG wire#powerrail
      "Order_Table_FB_Carousel_DB"(System_Selected := wire#w1, AutoMan_Switch := wire#w2, CurrentTime := "Time".CurrentLocalTime, CurrentDTL := "Time".CurrentDTL, Watchdog := "Watchdog_Settings", Cnv_Entry := "Control_DB".Inbound_Cnv, Cnv_PopUp_1 := "Control_DB".PopUp_Cnv[1], WeighingStation := "Weigh_Station_DB", ProfileStation := "Profile_Station_DB", Cnv_PopUp_2 := "Control_DB".PopUp_Cnv[2], Cnv_PopUp_3 := "Control_DB".PopUp_Cnv[3], Cnv_PopUp_4 := "Control_DB".PopUp_Cnv[4], Cnv_Exit := "Control_DB".Outbound_Cnv, System := "System_DB_Carousel", Control_OPC_Ua := "Control_DB"."Carrousel_Order Table")
   END_RUNG
   RUNG wire#powerrail
      Contact( "AlwaysTRUE" )
   END_RUNG wire#w1
   RUNG wire#powerrail
      Contact( "AlwaysTRUE" )
   END_RUNG wire#w2
   // the same network as SCL:
   "Order_Table_FB_Carousel_DB"(System_Selected := "AlwaysTRUE",   // "Order_Table_FB_Carousel"
                           AutoMan_Switch := "AlwaysTRUE",
                           CurrentTime := "Time".CurrentLocalTime,
                           CurrentDTL := "Time".CurrentDTL,
                           Watchdog := "Watchdog_Settings",
                           Cnv_Entry := "Control_DB".Inbound_Cnv,
                           Cnv_PopUp_1 := "Control_DB".PopUp_Cnv[1],
                           WeighingStation := "Weigh_Station_DB",
                           ProfileStation := "Profile_Station_DB",
                           Cnv_PopUp_2 := "Control_DB".PopUp_Cnv[2],
                           Cnv_PopUp_3 := "Control_DB".PopUp_Cnv[3],
                           Cnv_PopUp_4 := "Control_DB".PopUp_Cnv[4],
                           Cnv_Exit := "Control_DB".Outbound_Cnv,
                           System := "System_DB_Carousel",
                           Control_OPC_Ua := "Control_DB"."Carrousel_Order Table");
END_REGION

REGION Network 20: System Order Table - VTD and Conveyors
   RUNG wire#powerrail
      "Order_Table_FB_VTD_DB"(AutoMan_Switch := wire#w1, System_Selected := "AlwaysTRUE", CurrentTime := "Time".CurrentLocalTime, CurrentDTL := "Time".CurrentDTL, Watchdog := "Watchdog_Settings", VTD := "Control_DB".VTD_Control, Extrator_Conveyor := "Control_DB".ECnv_Control, Cnv_Buffer_1 := "Control_DB".LCnv_Control[1], Cnv_Buffer_2 := "Control_DB".LCnv_Control[2], Cnv_Buffer_3 := "Control_DB".LCnv_Control[3], System := "System_DB_VTD", Control_OPC_Ua := "Control_DB"."VTD_Order Table")
   END_RUNG
   RUNG wire#powerrail
      Contact( "AlwaysTRUE" )
   END_RUNG wire#w1
   // the same network as SCL:
   "Order_Table_FB_VTD_DB"(System_Selected := "AlwaysTRUE",   // "Order_Table_FB_VTD"
                           AutoMan_Switch := "AlwaysTRUE",
                           CurrentTime := "Time".CurrentLocalTime,
                           CurrentDTL := "Time".CurrentDTL,
                           Watchdog := "Watchdog_Settings",
                           VTD := "Control_DB".VTD_Control,
                           Extrator_Conveyor := "Control_DB".ECnv_Control,
                           Cnv_Buffer_1 := "Control_DB".LCnv_Control[1],
                           Cnv_Buffer_2 := "Control_DB".LCnv_Control[2],
                           Cnv_Buffer_3 := "Control_DB".LCnv_Control[3],
                           System := "System_DB_VTD",
                           Control_OPC_Ua := "Control_DB"."VTD_Order Table");
END_REGION

REGION Network 21: CLOCK AND HEARTBEATING *
   RUNG wire#powerrail
      "FC_CLOCK"(Ret_Val => "Time".CurrentDTL, CurrentTime => "Time".CurrentLocalTime)
      "FB_HeartBeat_DB"(PC_HeartBeat := "Time".PC_HeartBeat, PLC_HeartBeat => "Time".PLC_HeartBeat, PC_Disconnected =>)
   END_RUNG
   // the same network as SCL:
   "Time".CurrentDTL := "FC_CLOCK"(CurrentTime => "Time".CurrentLocalTime, ENO => #_w1);
   IF #_w1 THEN
       "FB_HeartBeat_DB"(PC_HeartBeat := "Time".PC_HeartBeat, PLC_HeartBeat => "Time".PLC_HeartBeat);   // "FB_HeartBeat"
   END_IF;
END_REGION
END_ORGANIZATION_BLOCK
